(* IEC 61131-3 sources: plc-process-lib/tools/demo/src/POUs/F_DemoEvent, 2 files *)

(* ---- F_DemoEvent.decl.st ---- *)
// Назначение: запись события сценария (действие «оператора», возмущение) в журнал событий
//             GVL_DemoLog для подписей на графиках. Журнал полон — событие не пишется, FALSE.
// Автор:      kr0nsch
// Версия:     0.1.0
// Документ:   docs/media/data/demo-events.csv; tools/demo/README.md
FUNCTION F_DemoEvent : BOOL
VAR_INPUT
    lrT_s     : LREAL;   // время события от старта сценария, с
    iScenario : INT;     // номер сценария: 1 — A, 2 — B, 3 — C
    iCode     : INT;     // код события (по сценарию)
END_VAR

(* ---- F_DemoEvent.impl.st ---- *)
IF GVL_DemoLog.uiEvN < GVL_DemoConst.EVENT_LOG_N THEN
    GVL_DemoLog.arEvT_s[GVL_DemoLog.uiEvN] := LREAL_TO_REAL(lrT_s);
    GVL_DemoLog.aiEvScenario[GVL_DemoLog.uiEvN] := iScenario;
    GVL_DemoLog.aiEvCode[GVL_DemoLog.uiEvN] := iCode;
    GVL_DemoLog.uiEvN := GVL_DemoLog.uiEvN + 1;
    F_DemoEvent := TRUE;
END_IF
